TYPE ST_FixtureRecord :
STRUCT
	nId : UDINT;
	fValue : LREAL;
	sLabel : STRING(40);
	eMode : E_FixtureMode;
END_STRUCT
END_TYPE

(* stored: Version 1.1.0.1
   DUT ST_FixtureRecord: Id {7253c2e2-06b0-4455-8b6b-2a9ddef35223} *)
